PROGRAM PLC_PRG
VAR
END_VAR

END_PROGRAM

(* stored: Version 1.1.0.1, ProductVersion 3.1.4024.16
   POU PLC_PRG: Id {ed5d9213-db5c-4467-b81d-16800f5128fe}, SpecialFunc None *)
